// TIA Portal V20 export
// export: Created 2026-10-20T18:54:42.1772018Z, ExportSetting None, DisplayName Totally Integrated Automation Portal, DisplayVersion V20 Update 6, DisplayName TIA Portal Openness, DisplayVersion V20 Update 6, DisplayName TIA Portal Version Control Interface, DisplayVersion V20 Update 6, DisplayName SINAMICS Startdrive Advanced, DisplayVersion V20 SP1, DisplayName SINAMICS Startdrive G130, G150, S120, S150, SINAMICS MV, G220, S200, S210, DisplayVersion V20 SP1, DisplayName SINAMICS Startdrive G110M, G120, G120C, G120D, G120P, G115D, DisplayVersion V20 SP1, DisplayName STEP 7 Professional, DisplayVersion V20 Update 6, DisplayName STEP 7 Safety, DisplayVersion V20 Update 2, DisplayName WinCC Basic/Comfort/Advanced, DisplayVersion V20 Update 6, DisplayName WinCC Unified, DisplayVersion V20 Update 6
VAR_GLOBAL   // PLC tag table "IO_Turck_1"
   "Light_Rear_1_Bounce_Style(1)" AT %QB159 : Byte;   // Last byte - 14
   "Light_Front_1_Pulse_Pattern(1)" AT %QB133 : Byte;   // Last byte - 8
   "Light_Rear_1_Pulse_Pattern(1)" AT %QB165 : Byte;   // Last byte - 8
   "Light_Rear_1_Color1(1)" AT %QB171 : Byte;   // Last byte - 2
   "Light_Front_1_Color1(1)" AT %QB139 : Byte;   // Last byte - 2
   "Light_Rear_1_Intensity2(1)" AT %QB161 : Byte;   // Last byte - 12
   "Light_Rear_1_Direction(1)" AT %QB147 : Byte;   // Last byte - 18
   "Light_Rear_1_Speed(1)" AT %QB167 : Byte;   // Last byte - 6
   "Light_Rear_1_Intensity1(1)" AT %QB169 : Byte;   // Last byte - 4
   "Light_Front_1_Intensity1(1)" AT %QB137 : Byte;   // Last byte - 4
   "Light_Front_1_Animation(1)" AT %QB141 : Byte;   // Last byte
   "Light_Front_1_Color2(1)" AT %QB131 : Byte;   // Last byte - 10
   "Light_Rear_1_Percent_Width1(1)" AT %QB157 : Byte;   // Last byte - 16
   "Light_Front_1_Percent_Width1(1)" AT %QB125 : Byte;   // Last byte - 16
   "Light_Front_1_Intensity2(1)" AT %QB129 : Byte;   // Last byte - 12
   "Light_Front_1_Bounce_Style(1)" AT %QB127 : Byte;   // Last byte - 14
   "Light_Rear_1_Animation(1)" AT %QB173 : Byte;   // Last byte
   "Light_Front_1_Speed(1)" AT %QB135 : Byte;   // Last byte - 6
   "Light_Rear_1_Color2(1)" AT %QB163 : Byte;   // Last byte - 10
   "Light_Front_1_Direction(1)" AT %QB123 : Byte;   // Last byte - 18
END_VAR
